Staubli VAL3: setAlarm.pgx

public program setAlarm(num x_nAlarmCode (dimensions=1), num x_nErrIndex (dimensions=1))
  local bool l_bExist
  local num l_nIndex
  local string l_sAlarmLevel
  local string l_sErrMsg
begin
  //check if the alarm has existed in the list
  do
    l_bExist=(x_nAlarmCode==_nAlarmCode[l_nIndex] and x_nErrIndex==_nErrIndex[l_nIndex])
    l_nIndex=l_nIndex+1
  until l_bExist or l_nIndex>=size(_nAlarmCode)
  //
  if !l_bExist
    //new alarm, add it
    if _nAlarmCode[_nAlarmIndex]>0
      _nAlarmIndex=(_nAlarmIndex+1)%size(_nAlarmCode)
    endIf
    _nAlarmCode[_nAlarmIndex]=x_nAlarmCode
    _nErrIndex[_nAlarmIndex]=x_nErrIndex
    call getAlarmMsg(x_nAlarmCode,l_sErrMsg)
    //错误等级
    if _nAlarmCode[_nAlarmIndex]>=0
      if x_nAlarmCode>nHeavyAlarmLev
        l_sAlarmLevel="错误："
      else
        l_sAlarmLevel="警告："
      endIf
      //错误消息
      if x_nErrIndex>=0
        sAlarmMes[_nAlarmIndex]=_sRobotStatus=l_sAlarmLevel+"-"+toString("",x_nAlarmCode)+". "+":"+toString("",x_nErrIndex)+l_sErrMsg
      else
        sAlarmMes[_nAlarmIndex]=_sRobotStatus=l_sAlarmLevel+"-"+toString("",x_nAlarmCode)+". "+l_sErrMsg
      endIf
      logMsg(sAlarmMes[_nAlarmIndex])
    endIf
    delay(0)
  endIf
end
